(*
SPDX-FileCopyrightText: © 2026 Oleksandr Tiutyk <trofimich@gmail.com>
SPDX-License-Identifier: MIT
License: https://opensource.org/license/mit
*)

(*!
<summary>Checks the configured new interval after late start-preparation refusal.</summary>
<description>
The case executes in one PLC callback with a persistent restart probe and no external resources.
AfterTest prepares the fixture for reuse by the runner.
</description>
*)

{attribute 'no_assign'}
{attribute 'no_explicit_call' := 'do not call this function block directly'}
FUNCTION_BLOCK TimerRestartStartFailureTest EXTENDS TOF_Testing.SingleCycleTest
VAR_STAT
	{attribute 'hide'}
	_ClassName : STRING := __POUNAME();
END_VAR
VAR CONSTANT
	//! <summary>Positive interval selected for the replacement run.</summary>
	_PositiveInterval : TIME := T#30MS;
END_VAR
VAR
	_Timer : TimerRestartProbe(name := "Start refusal");
END_VAR

(*!
<summary>Checks the configured new interval after late start-preparation refusal.</summary>
*)
METHOD PROTECTED ExecuteTest
_Timer.Interval := TOF_Core.Times.MIN_VALUE;
_Timer.ThrowOnBeforeStart := TRUE;
Assert.ThatBool(
	actual := _Timer.SetIntervalAndRestart(interval := _PositiveInterval),
	message := "Start preparation exception must be converted to restart refusal"
).IsFalse();
Assert.ThatBool(
	actual := _Timer.State.Ready,
	message := "Refused Start must leave the prepared timer READY"
).IsTrue();
Assert.ThatBool(
	actual := _Timer.Interval = _PositiveInterval,
	message := "Late Start refusal must retain the new PT"
).IsTrue();
Assert.ThatBool(
	actual := _Timer.Elapsed,
	message := "Injected refusal before base Start must leave Q clear"
).IsFalse();
_Timer.Execute();
Assert.ThatBool(
	actual := _Timer.State.Ready,
	message := "Refused restart must not schedule automatic execution"
).IsTrue();
_Timer.ThrowOnBeforeStart := FALSE;

IF NOT _Timer.Start() THEN
	RecordFailure(message := "Explicit Start must recover after removing injection");
	RETURN;
END_IF

IF NOT _Timer.Cancel() THEN
	RecordFailure(message := "Scenario must cancel the recovered run");
	RETURN;
END_IF

_Timer.Execute();
Assert.ThatBool(
	actual := _Timer.State.Stopped AND_THEN _Timer.FinalStopReason.ExternalCancel,
	message := "The replacement run must finish cancellation"
).IsTrue();
END_METHOD

(*!
<summary>Returns the owned timer to READY before reporting the result.</summary>
<description>
Reopens the stopping gate and disables callback injections before cooperative cleanup.
</description>
*)
METHOD PROTECTED AfterTest
_Timer.AllowStopping := TRUE;
_Timer.ThrowOnBeforeStart := FALSE;
_Timer.ThrowOnReset := FALSE;
_Timer.ResetOnAfterStop := FALSE;

Assert.ThatBool(
	actual := PrepareTimerTestForReuse(timer := _Timer),
	message := "The timer must return to READY after cleanup"
).IsTrue();
END_METHOD

//! <summary>Borrows the concrete class name. Callers must not modify it.</summary>
{attribute 'monitoring' := 'call'}
PROPERTY ClassName : REFERENCE TO STRING
GET
ClassName REF= _ClassName;
END_GET
END_PROPERTY

//! <summary>Borrows the compiler-initialized namespace. Callers must not modify it.</summary>
{attribute 'monitoring' := 'call'}
PROPERTY NamespaceName : REFERENCE TO STRING
GET
NamespaceName REF= CurrentNamespace.Name;
END_GET
END_PROPERTY

//! <summary>Reports the concrete instance size in bytes.</summary>
{attribute 'monitoring' := 'call'}
PROPERTY SelfSize : ULINT
GET
SelfSize := XSIZEOF(THIS^);
END_GET
END_PROPERTY

END_FUNCTION_BLOCK

(* stored: Version 1.1.0.1
   POU TimerRestartStartFailureTest: Id {071ea9cf-9816-4eb6-bcb2-055b98bd213f}, SpecialFunc None
   Method ExecuteTest: Id {275c69cd-cdc0-4dd3-b766-3a22e55f88f3}
   Method AfterTest: Id {51c7d455-2c88-47a0-a8c7-b24bb0aa3b16}
   Property ClassName: Id {234cc419-1cac-43c4-aa6b-399e2540c426}
   Get Get: Id {48568fa1-9c3a-4fe6-9ff4-a31453b23343}
   Property NamespaceName: Id {8bd275dc-2c57-40d9-ad23-4db742bcd62d}
   Get Get: Id {545a43c2-b6cc-4a2e-98d4-782cdfe516f4}
   Property SelfSize: Id {11587047-1490-464b-9858-664106eeabd7}
   Get Get: Id {5b9dca2f-a4d5-4a0c-ae3e-5cfb5c1c0c27} *)
